(* IEC 61131-3 sources: llm-plc-st-eval/data/processed_v2/gpt-4o/I2/zero_shot, 3 files *)

(* ---- ejec_1.st ---- *)
FUNCTION_BLOCK FB_Llenado
VAR
    // Entradas
    nivelAlto : BOOL;    // Sensor de nivel alto
    nivelBajo : BOOL;    // Sensor de nivel bajo
    btnInicio : BOOL;    // Botón de inicio
    btnParo : BOOL;      // Botón de paro

    // Salidas
    vLlenado : BOOL;     // Válvula de llenado
    motorMezcla : BOOL;  // Motor de mezcla
    vDescarga : BOOL;    // Válvula de descarga

    // Variables internas
    estado : INT;        // Estado del proceso
    timerMezcla : TON;   // Temporizador para el motor de mezcla
END_VAR

// Inicialización del bloque de función
IF NOT btnParo THEN
    CASE estado OF
        0: // Estado de reposo
            vLlenado := FALSE;
            motorMezcla := FALSE;
            vDescarga := FALSE;
            IF btnInicio THEN
                estado := 1; // Ir al estado de llenado
            END_IF;

        1: // Estado de llenado
            vLlenado := TRUE;
            IF nivelAlto THEN
                vLlenado := FALSE;
                estado := 2; // Ir al estado de mezcla
                timerMezcla(IN := TRUE, PT := T#60S);
            END_IF;

        2: // Estado de mezcla
            motorMezcla := TRUE;
            timerMezcla(IN := TRUE);
            IF timerMezcla.Q THEN
                motorMezcla := FALSE;
                estado := 3; // Ir al estado de descarga
            END_IF;

        3: // Estado de descarga
            vDescarga := TRUE;
            IF nivelBajo THEN
                vDescarga := FALSE;
                estado := 0; // Volver al estado de reposo
            END_IF;
    END_CASE;
ELSE
    // Estado seguro en caso de paro
    vLlenado := FALSE;
    motorMezcla := FALSE;
    vDescarga := FALSE;
    estado := 0; // Volver al estado de reposo
    timerMezcla(IN := FALSE);
END_IF;
END_FUNCTION_BLOCK

(* ---- ejec_2.st ---- *)
FUNCTION_BLOCK FB_Llenado
VAR
    // Entradas
    nivelAlto : BOOL;
    nivelBajo : BOOL;
    btnInicio : BOOL;
    btnParo : BOOL;

    // Salidas
    vLlenado : BOOL := FALSE;
    motorMezcla : BOOL := FALSE;
    vDescarga : BOOL := FALSE;

    // Variables internas
    estado : INT := 0; // 0: Reposo, 1: Llenado, 2: Mezcla, 3: Descarga
    timerMezcla : TON; // Temporizador para el motor de mezcla
END_VAR

// Inicialización del temporizador
timerMezcla(IN := FALSE, PT := T#60S);

IF btnParo THEN
    // Si se presiona el botón de paro, se desactivan todas las salidas y se vuelve a reposo
    vLlenado := FALSE;
    motorMezcla := FALSE;
    vDescarga := FALSE;
    estado := 0;
ELSE
    CASE estado OF
        0: // Reposo
            IF btnInicio THEN
                estado := 1; // Cambiar al estado de llenado
            END_IF;

        1: // Llenado
            vLlenado := TRUE;
            IF nivelAlto THEN
                vLlenado := FALSE;
                estado := 2; // Cambiar al estado de mezcla
                timerMezcla(IN := TRUE); // Iniciar temporizador de mezcla
            END_IF;

        2: // Mezcla
            motorMezcla := TRUE;
            timerMezcla(IN := TRUE);
            IF timerMezcla.Q THEN
                motorMezcla := FALSE;
                estado := 3; // Cambiar al estado de descarga
            END_IF;

        3: // Descarga
            vDescarga := TRUE;
            IF nivelBajo THEN
                vDescarga := FALSE;
                estado := 0; // Volver al estado de reposo
            END_IF;
    END_CASE;
END_IF;
END_FUNCTION_BLOCK

(* ---- ejec_3.st ---- *)
FUNCTION_BLOCK FB_Llenado
VAR
    // Variables de entrada
    nivelAlto : BOOL;    // Sensor de nivel alto
    nivelBajo : BOOL;    // Sensor de nivel bajo
    btnInicio : BOOL;    // Botón de inicio
    btnParo   : BOOL;    // Botón de paro

    // Variables de salida
    vLlenado    : BOOL;  // Válvula de llenado
    motorMezcla : BOOL;  // Motor de mezcla
    vDescarga   : BOOL;  // Válvula de descarga

    // Variables internas
    estado      : INT;   // Estado del proceso
    timerMezcla : TON;   // Temporizador para el motor de mezcla
END_VAR

// Inicialización del temporizador
timerMezcla(IN := FALSE, PT := T#60S);

// Lógica del proceso de llenado por etapas
IF btnParo THEN
    // Si se presiona el botón de paro, llevar todo a estado seguro
    estado := 0;
    vLlenado := FALSE;
    motorMezcla := FALSE;
    vDescarga := FALSE;
ELSIF btnInicio THEN
    CASE estado OF
        0: // Estado de reposo
            IF btnInicio THEN
                estado := 1; // Iniciar proceso de llenado
            END_IF;

        1: // Estado de llenado
            vLlenado := TRUE;
            IF nivelAlto THEN
                vLlenado := FALSE;
                estado := 2; // Pasar al estado de mezcla
            END_IF;

        2: // Estado de mezcla
            motorMezcla := TRUE;
            timerMezcla(IN := TRUE);
            IF timerMezcla.Q THEN
                motorMezcla := FALSE;
                timerMezcla(IN := FALSE);
                estado := 3; // Pasar al estado de descarga
            END_IF;

        3: // Estado de descarga
            vDescarga := TRUE;
            IF nivelBajo THEN
                vDescarga := FALSE;
                estado := 0; // Volver al estado de reposo
            END_IF;
    END_CASE;
END_IF;
END_FUNCTION_BLOCK
